  global container_id = 0
  global powder_id  = 0
  global bulk_density = 0
  global H          = 0
  global H_c          = 0
  global mouth_d     = 0
  global mouth_sh    = 0
  global length_c     = 0
  global diameter   = 0
  global empty_weight_g  = 0
  global volume_ml    = 0
  global shape_code   = 0
  global flow_code   = 0
  global shape = ""
  global Flowability = ""
  global full_weight_g = 0
  global cent_edge = 0
  global pick_2_base = 0.2 # distance from tcp to base of picking table
  global wall_thickness = 0.002

  def read_db_data():

    socket_open(SERVER_IP, SERVER_PORT)
    sleep(0.5)
    socket_send_string("GET_DATACODE_FLOATS")
    sleep(5)

    local fl = socket_read_ascii_float(14)
    socket_close()

    global container_id = fl[1]
    global powder_id = fl[2]
    global bulk_density = fl[3]
    global H          = fl[4]/1000
    global H_c          = fl[5]/1000
    global mouth_d     = fl[6]/1000
    global mouth_sh    = fl[7]/1000
    global length_c     = fl[8]/1000
    global diameter   = fl[9]/1000
    global empty_weight_g = fl[10]
    global volume_ml    = fl[11]
    global full_weight_g = fl[12]
    global flow_code   = fl[13]
    global shape_code   = fl[14]

  	if (flow_code == 1.0):
  	  global Flowability = "MEDIUM"
  	elif (flow_code == 2.0):
  	  global Flowability = "LOW"
  	else:
  	  global Flowability = "HIGH"
  	end

    if ( shape_code == 1.0):
  	shape = "cylindrical"
  	cent_edge =  diameter
    else:
  	shape = "cubical"
  	cent_edge =  length_c
    end

  end

  def send_picking_info(Pow_name, target_weight):
    socket_open(SERVER_IP, SERVER_PORT)
    cmd = "PICK:"+Pow_name+";"+to_str(target_weight)
    socket_send_string(cmd)
    sleep(0.1)
    socket_close()
  end

  #### POTS ####
  def tilt_send(angle):
  	socket_open(SERVER_IP, SERVER_PORT)
  	angle = 92.0 - angle
  	socket_send_string("TILT:"+to_str(angle))
  	sync()
  	sleep(0.5)
  	socket_close()
  end

  def CW_Rotate(angle):
  	socket_open(SERVER_IP, SERVER_PORT)
  	socket_send_string("CWROTATE:"+to_str(angle))
  	sync()
  	sleep(0.5)
  	socket_close()
  end

  def CCW_Rotate(angle):
  	socket_open(SERVER_IP, SERVER_PORT)
  	socket_send_string("CCWROTATE:"+to_str(angle))
  	sync()
  	sleep(0.5)
  	socket_close()
  end

  def CW_full_Rotate():
  	socket_open(SERVER_IP, SERVER_PORT)
  	socket_send_string("FULLROTATE:"+to_str(1))
  	sync()
  	sleep(0.5)
  	socket_close()
  end

  def CCW_full_Rotate():
  	socket_open(SERVER_IP, SERVER_PORT)
  	socket_send_string("FULLROTATE:"+to_str(-1))
  	sync()
  	sleep(0.5)
  	socket_close()
  end

  def tilt_to_home():
  	socket_open(SERVER_IP, SERVER_PORT)
  	socket_send_string("HOME")
  	sync()
  	sleep(0.5)
  	socket_close()
  end
  #######
  def vibration_1():
  	set_analog_out(0,0.4)
  	sleep(1)
  	set_analog_out(0,0.0)
  	sleep(0)
  end

  def vibration_2():
  	set_analog_out(0,0.4)
  	sleep(0.8)
  	set_analog_out(0,0.0)
  	sleep(0.2)
  end

  def vibration_3():
  	set_analog_out(0,0.4)
  	sleep(0.5)
  	set_analog_out(0,0.0)
  	sleep(0.3)
  end

  def vibration_4():
  	set_analog_out(0,0.4)
  	sleep(0.5)
  	set_analog_out(0, 0.0)
  	sleep(0.5)
  end

  def vibration_5():
  	set_analog_out(0,0.4)
  	sleep(0.2)
  	set_analog_out(0, 0.0)
  	sleep(0.8)
  end

  ##################

  global gear_2_holder = 0.018
  global gain_per_percent = 0.5
  global hinge_2_base = 0.0421
  global TCP_2_tip_x = 0.0047
  global spatula_len = 0.182
  global spatula_offset = p[TCP_2_tip_x,0,spatula_len,0,0,0]
  global SPATULA_L_VOL_ML = 5.0        # 1 teaspoon = 5 mL
  global SPATULA_M_VOL_ML = 1.25       # 1/4 teaspoon = 1.25 mL
  global SPATULA_S_VOL_ML = 0.15625    # 1/32 teaspoon = 0.15625 mL
  global SPATULA_FLAT_M_VOL_ML  = 2.2
  global SPATULA_FLAT_S_VOL_ML  = 0.7   #based on caluclations using rho = m/V

  def correction_reset():
  	global g_k = 0.0
  	global g_depth_corr = 0.0
  	global g_prev_cum_w = weight_value
  end

  def params_init():

  	global scoop_status= ""
  	global w_dosed_total = 0.0
  	global last_scale = 0.0
  	global tilt_angle_sent = 0.0
  	global level = 0.0
  	global target_g = 0.0
  	global angle_max = 70
  	global angle_min = 20
  	global ry_deg_safe = 0
  	global ry_deg = 0

  	global scoop_ct = 0
  	global error_sum = 0.0
  	global error_sq_sum = 0.0
  	global scoop_g = 0.0

  	global g_k =0.0
  	global g_eta = 0.3

  	global g_gain_scale = 0.07
  	global g_k_min = 0.0
  	global g_k_max = 0.09

  	# ---------- Damping ----------
  	global g_alpha_under = 0.75   # aggressive when undershooting
  	global g_alpha_over  = 0.30   # conservative when overshooting

  	# ---------- Search ----------
  	global g_engagement_min = 0.05
  	global g_search_step = 0.01      # 3 mm

  	# ---------- Deadband ----------
  	global g_tol = 0.02               # 20 mg minimum
  	global g_tol_ratio = 0.05         # ±5% of target

  	# ---------- Limits ----------
  	global g_corr_max = 0.020         # 20 mm maximum correction

  	# ---------- States ----------
  	global g_depth_corr = 0.0
  	global g_prev_cum_w = -1.0
  end

  def clamp(x, lo, hi):
  	if(x<lo):
  		return lo
  	elif (x>hi):
  		return hi
  	else:
  		return x
  	end
  end

  def compute_level_percent(W_now, weight_value):   # W_now = container+powder, weight_value = live scale reading
      global delta = weight_value - last_scale

      if (delta < 0.0):
          delta = 0.0
      end

      global w_dosed_total = w_dosed_total + delta
      global last_scale = weight_value     # update the last scale reading

      local W_eff = W_now - w_dosed_total
      if (W_eff <  empty_weight_g):
          W_eff =  empty_weight_g
      end

      # Compute powder level %
      level = 100.0 * (W_eff -  empty_weight_g) / (full_weight_g -  empty_weight_g)

      # Clamp to 0–100
      level = clamp(level, 0, 100)
    textmsg("deb 1 = ", level)
      return level
  end

  def deg2rad(d):
  	return d*3.141592/180
  end

  def my_abs(val):
  	if (val<0):
  		return -val
  	else:
  		return val
  	end
  end

  def compute_tilt_deg(level_percent):
  	angle = angle_min + gain_per_percent*(100.0-level_percent)

    	textmsg("deb 2 = ", angle)
  	return clamp(angle, angle_min, angle_max)
  end

  def tilt(level_percentage):
  	new_angle = compute_tilt_deg(level_percentage)
    	textmsg("deb angle 1 = ", new_angle)
  	global angle_rel = new_angle - tilt_angle_sent
    	textmsg("deb 2 = ", angle_rel)

  	if my_abs(angle_rel)>2.0:
    		textmsg("deb loop")
  		tilt_send(new_angle)
  		global angle_deg = new_angle
    		textmsg("deb 2 = ", angle_deg)
  		global tilt_angle_sent = new_angle
  		global p_center_vertical = center_pose()
  		global p_center = updated_center_pose(p_center_vertical, angle_deg)
  	end
    	textmsg("deb loop exit")

  	tilt_send(angle_deg)
    	textmsg("deb angle 2 =", angle_deg)

  end

  def compute_scoop_depth(level, weight_value, target_g):

      global scoop_depth_rel = ((100.0-level)/100.0)*(H-mouth_sh)

      if (g_prev_cum_w < 0):
          g_prev_cum_w = weight_value
          g_depth_corr = 0.0

      else:
          global scoop_g = weight_value - g_prev_cum_w
          g_prev_cum_w = weight_value

          local error = target_g - scoop_g
          local engagement = scoop_g / target_g

          local tol = g_tol_ratio * target_g
          if (tol < g_tol):
              tol = g_tol
          end
          if ((engagement < g_engagement_min) and (scoop_g < target_g)):
              g_depth_corr = g_depth_corr + g_search_step
          elif (my_abs(error) <= tol):
  			sync()
          else:
              local error_norm = my_abs(error / target_g)
              local g_target = clamp(g_gain_scale * error_norm,g_k_min,g_k_max)

              g_k = (1.0-g_eta) * g_k + g_eta * g_target
              if (error > 0):
                  local corr = g_k * error
                  g_depth_corr = g_depth_corr +g_alpha_under * corr
              else:
                  local corr = g_k * error
                  g_depth_corr = g_depth_corr +g_alpha_over * corr

              end
              g_depth_corr = clamp(g_depth_corr,-g_corr_max,g_corr_max)

          end
      end
      scoop_depth = scoop_depth_rel + g_depth_corr
      scoop_depth = clamp(scoop_depth, 0.0, H)
      return scoop_depth

  end

  def get_scoop_weight(spatula, bulk_density):

  	local vol = 0

  	if (spatula == "spatula_L"):
  		vol = SPATULA_L_VOL_ML
  		global spatula_depth = 0.015
  		global spatula_mid   = 0.016
  		global spatula_ry    = 0.0

  	elif (spatula == "spatula_M"):
  		vol = SPATULA_M_VOL_ML
  		global spatula_depth = 0.010
  		global spatula_mid   = 0.0105
  		global spatula_ry    = 0.0

  	elif (spatula == "spatula_S"):
  		vol = SPATULA_S_VOL_ML
  		global spatula_depth = 0.008
  		global spatula_mid   = 0.006
  		global spatula_ry    = 0.0

  	elif (spatula == "spatula_flat_M"):
  		vol = SPATULA_FLAT_M_VOL_ML
  		global spatula_depth = 0.005
  		global spatula_mid   = 0.02
  		global spatula_ry    = 4.0

  	elif (spatula == "spatula_flat_S"):
  		vol = SPATULA_FLAT_S_VOL_ML
  		global spatula_depth = 0.005
  		global spatula_mid   = 0.011
  		global spatula_ry    = 4.0
  	else:
  		textmsg("Unknown spatula type")
  		return 0.0
  	end
  	global target_g = vol * bulk_density
  	return target_g

  end

  def select_spatula(Flowability, level, diff, bulk_density, mouth_d ):

      local k = 1.1
      global powder_height = (H  - mouth_sh ) * level/100

      if (Flowability == "LOW"):
          local gFM = get_scoop_weight("spatula_flat_M", bulk_density)
  		local level_ok_FM = (mouth_d >= 0.05)
          local level_ok_FM = (spatula_mid  < powder_height)
          local diff_ok_FM  = (diff > k * gFM)
          local flatM_ok = level_ok_FM and diff_ok_FM
          if (flatM_ok):
              return "spatula_flat_M"
          else:
              return "spatula_flat_S"
          end
      end

      local gL = get_scoop_weight("spatula_L", bulk_density)
      local mouth_ok_L = (mouth_d  >= 0.05)
      local level_ok_L = (spatula_mid < powder_height)
      local diff_ok_L  = (diff > k * gL)

      local large_ok = mouth_ok_L and level_ok_L and diff_ok_L
      local gM = get_scoop_weight("spatula_M", bulk_density)
      local level_ok_M = (spatula_mid < powder_height)
      local diff_ok_M  = (diff > k * gM)

      local medium_ok = level_ok_M and diff_ok_M

      if (large_ok):
          return "spatula_L"
      elif (medium_ok):
          return "spatula_M"
      else:
          return "spatula_S"
      end
  end

  def after_scoop():
  	set_tcp(tcp_dosing)
  	set_analog_out(0,0.0)
  	tilt_send(angle_deg)
  	sleep(0.5)
  	movel(lifted_pose, a=0.05, v=0.2)
  	movel(tilted_pose_in_base2, a=0.05, v=0.2)
  	set_analog_out(0,0.4)
  	if (Flowability == "LOW"):
  		movel(end_rel_tilted_level2, a=0.03, v=0.1)
  		sleep(0.5)
  		movel(tilted_pose_in_base2, a=0.05, v=0.2)
  	  	movel(pose_trans(tilted_pose_in_base2, p[0,0,0,0,0,2.0]), a=0.05, v=0.2)
  		#movel(tilted_pose_in_base2, a=0.05, v=0.2)
  	else:
  	    movel(pose_trans(tilted_pose_in_base2, p[0,0,0,0,0,2.0]), a=0.05, v=0.2)
  	    movel(tilted_pose_in_base2, a=0.05, v=0.2)
  	end
  	set_analog_out(0,0.0)
  	movel(lifted_pose, a=0.5, v=0.5)
  	tilt_to_home()
  	set_tcp(tcp_default)
  end

  def center_pose():
  	global p_translated = container_place
  	#global p_translated = pots_axis_temp

  	#cx = p_translated[0]
  	#cy = p_translated[1]
  	#cz = p_translated[2]

  	global p_center_vertical_temp = pose_trans(p_translated, p[0,0,0, deg2rad(90), 0, 0])
  	cx = p_center_vertical_temp[0]
  	cy = p_center_vertical_temp[1]
  	cz = p_center_vertical_temp[2]
  	rx = p_center_vertical_temp[3]
  	ry = p_center_vertical_temp[4]
  	rz = p_center_vertical_temp[5]

  	global p_center_vertical_temp = p[cx,cy,cz, 0, 0, rz]
  	trans_rel = p[0,0,-pick_2_base+H,0,0,0]
  	global p_center_vertical =  pose_trans(p_center_vertical_temp, trans_rel)
  	return p_center_vertical
  end

  def updated_center_pose(p_center_vertical, angle_deg):
  	hinge_pose = pose_trans(p_center_vertical, p[0,0,-hinge_2_base-gear_2_holder-H ,0,0,0])
  	local_rel = pose_trans(pose_inv(hinge_pose), p_center_vertical)

  	rot_tilt = p[0,0,0, -deg2rad(angle_deg),0,0]
  	local_rel_tilted = pose_trans(rot_tilt, local_rel)

  	global p_center = pose_trans(hinge_pose, local_rel_tilted)
  	return p_center
  end

  def scoop_powder(p_center):
  	vibration_voltage = 0.4
  	global scoop_radius_default = 0.0

  	scoop_radius_default = mouth_d /2 - spatula_depth - wall_thickness
  	scoop_safe_entry_pose = pose_trans(p_center, p[-TCP_2_tip_x,0,spatula_len+0.05,0,0,0])
  	scoop_entry_pose = pose_trans(p_center, p[-TCP_2_tip_x,0,spatula_len,0,0,0])

  	movel(scoop_safe_entry_pose, a=0.1, v=0.25)
  	movel(scoop_entry_pose, a=0.1, v=0.25)

  	scoop_start_rel_int = p[0, 0, -mouth_sh , 0, 0, 0]
  	scoop_start_pose_int = pose_trans(scoop_entry_pose, scoop_start_rel_int)


  	#local ry_deg = map_tilt_to_ry_deg(angle_deg,level)
  	#local ry_result = map_tilt_to_ry_deg(angle_deg,level)

  	#global scoop_depth = compute_scoop_depth(level,weight_value, target_g)

  	global ry = deg2rad(90-angle_deg)

  	#global ry_safe = ry_result[0]
  	#global ry = deg2rad(ry_result[1])

  	if (spatula_mid < powder_height):

  		global total_depth = mouth_sh + scoop_depth + spatula_mid
  		global total_depth = clamp(total_depth, 0, H - spatula_mid)

  		safe_scoop_pivot = (mouth_d  - spatula_depth)/(total_depth)
  		global ry_safe = asin(safe_scoop_pivot)

  		scoop_start_rel = p[scoop_radius_default, 0, -total_depth, 0, 0, 0]

  		rot_mid = p[0, 0, 0, 0, 0, 0.785]
  		rot_end = p[0, 0, 0, 0, 0, 1.5708]

  		scoop_via_rel = pose_trans(rot_mid, scoop_start_rel)
  		scoop_end_rel = pose_trans(rot_end, scoop_start_rel)

  		scoop_start_pose = pose_trans(scoop_entry_pose, scoop_start_rel)
  		scoop_via_pose = pose_trans(scoop_entry_pose, scoop_via_rel)
  		scoop_end_pose = pose_trans(scoop_entry_pose, scoop_end_rel)


  			if (Flowability == "LOW"):
  				movel(pose_trans(scoop_start_pose_int,p[0,0,0,0,0,-1.5708]), a=0.1, v=0.25)
  				local spatula_base = pose_trans(scoop_entry_pose, p[0, 0, -H+wall_thickness, 0, 0, 0])
  				local scrape_pivot = pose_trans(scoop_entry_pose, p[0,0, -spatula_len,0,0,0])

  				global sticky_in_angle = -atan((cent_edge/2-spatula_depth)/H)
  				spatula_tilt_rel = pose_trans(pose_inv(scrape_pivot), spatula_base)

  				spatula_tilt = pose_trans(spatula_tilt_rel, p[0, 0, 0, 0, sticky_in_angle, 0])
  				global tilted_pose = pose_trans(scrape_pivot, p[0,0,0,spatula_tilt[3],spatula_tilt[4], spatula_tilt[5]])

  				global tilted_pose = pose_trans(tilted_pose, p[0,0,spatula_len-H+wall_thickness,0,0,0])
  				global rotate_90=pose_trans(tilted_pose,p[0,0,0,0,0,-1.5708])


  				movel(rotate_90,a=0.1, v=0.25)

  				#global sticky_in_angle = -atan((cent_edge/2-wall_thickness-spatula_depth)/(total_depth+spatula_mid))
  				#local scrape_target = pose_trans(scoop_entry_pose, p[0,0,-total_depth-spatula_mid,0,0,0])
  				#local scrape_pivot = pose_trans(scoop_entry_pose, p[0,0,-spatula_len,0,0,0])
  				#local scrape_rel = pose_trans(pose_inv(scrape_pivot), scrape_target)
  				#local scoop_sticky_in = pose_trans(scrape_rel, p[0,0,0,0,sticky_in_angle,0])

  				#global scrape_pose = pose_trans(scrape_pivot, p[0,0,0,scoop_sticky_in[3],scoop_sticky_in[4], scoop_sticky_in[5]])
  				#global scrape_pose = pose_trans(scrape_pose, p[0,0,spatula_len-total_depth-spatula_mid,0,0,0])

  				#scoop_sticky_in = pose_trans(scoop_start_pose, p[0,0,0,0,sticky_in_angle,0])
  				#movel(scrape_pose, a=0.1, v=0.25)
  				#movel(scrape_target,a=0.1,v=0.25)
  				CW_full_Rotate()
  				movel(scoop_start_pose, a=0.1, v=0.25)

  			else:
  				movel(scoop_start_pose_int, a=0.1, v=0.25)
  				movel(scoop_start_pose, a=0.1, v=0.25)
  				CW_full_Rotate()
  			end

  		movec(scoop_via_pose, scoop_end_pose, a=0.05, v=0.04)
  		#sleep(1.0)

  		# safe_retention
  		local pivot_pose = pose_trans(scoop_end_pose, p[0,0,total_depth-spatula_len,0,0,0])
  		local end_rel = pose_trans(pose_inv(pivot_pose), scoop_end_pose)
  		local end_rel_tilted = pose_trans(end_rel, p[0, 0, 0, 0, ry_safe-deg2rad(spatula_ry), 0])
  		local tilted_pose_in_base = pose_trans(pivot_pose, p[0,0,0,end_rel_tilted[3],end_rel_tilted[4], end_rel_tilted[5]])
  		local tilted_pose_in_base = pose_trans(tilted_pose_in_base, p[0, 0, spatula_len-total_depth, 0, 0, 0])
  		# sptula pivoted around the container rim of the mouth at ry_safe
  		movel(tilted_pose_in_base, a=0.03, v=0.1)

  		global safe_x = sin(ry_safe)*(total_depth-mouth_sh - (mouth_d - spatula_depth)*tan(ry_safe/2))
  		global safe_z = cos(ry_safe)*(total_depth-mouth_sh - (mouth_d - spatula_depth)*tan(ry_safe/2))

  		local safe_up = pose_trans(tilted_pose_in_base, p[-safe_x,0,safe_z,0,0,0])
  		movel(safe_up, a=0.03, v=0.1)

  		# full exit
  		local pivot_pose2 = pose_trans(scoop_entry_pose, p[0,0,-spatula_len,0,0,0])
  		local end_rel2 = pose_trans(pose_inv(pivot_pose2), tilted_pose_in_base)
  		#popup("is the spatula crashing front? ", blocking = True)
  		local end_rel_tilted2 = pose_trans(end_rel2, p[0, 0, 0, 0, ry-ry_safe-deg2rad(spatula_ry), 0])

  	else : # emptying logic
  		CCW_full_Rotate()

  		spatula_base = pose_trans(scoop_entry_pose, p[0, 0, -H+wall_thickness, 0, 0, 0])
  		local pivot_pose2 = pose_trans(scoop_entry_pose, p[0,0,-spatula_len,0,0,0])
  		# tilt inwards
  		global in_angle = -atan((cent_edge/2-spatula_depth)/H)
  		spatula_tilt_rel = pose_trans(pose_inv(pivot_pose2), spatula_base)

  		spatula_tilt = pose_trans(spatula_tilt_rel, p[0, 0, 0, -in_angle, 0, 0])
  		global tilted_pose = pose_trans(pivot_pose2, p[0,0,0,spatula_tilt[3],spatula_tilt[4], spatula_tilt[5]])

  		global tilted_pose = pose_trans(tilted_pose, p[0,0,spatula_len-H+wall_thickness,0,0,0])

  		movel(tilted_pose,a=0.1, v=0.25)

  		rotate90=pose_trans(tilted_pose,p[0,0,0,0,0,1.5708])

  		#sleep(1)
  		#Rotate()
  		#sleep(0.2)
  		movel(rotate90, a=0.1, v=0.1)
  		#popup("is the spatula crashing front? ", blocking = True)
  		movel(pose_trans(scoop_start_pose_int,p[0,0,0,0,0,1.5708]), a=0.03, v=0.1)
  		# full exit
  		#local pivot_pose2 = pose_trans(scoop_entry_pose, p[0,0,-spatula_len,0,0,0])
  		local end_rel2 = pose_trans(pose_inv(scoop_entry_pose), rotate90)
  		local end_rel_tilted2 = pose_trans(end_rel2, p[0, 0, 0, 0, ry-in_angle-deg2rad(spatula_ry), 0])
  	end

  	# exit flat spoon
  	global tilted_pose_in_base2 = pose_trans(pivot_pose2, p[0,0,0,end_rel_tilted2[3],end_rel_tilted2[4], end_rel_tilted2[5]])
  	global tilted_pose_in_base2 = pose_trans(tilted_pose_in_base2, p[0, 0, spatula_len-spatula_mid, 0, 0, 0])
  	# spaula exited at center of the mouth at ry
  	movel(tilted_pose_in_base2, a=0.03, v=0.1)
  	if(scoop_status== "normal"):
  		vib_thread=True
  		if (spatula=="spatula_S"):
  			vibration_3()
  			local ry_level = deg2rad(12)
  		elif(spatula=="spatula_flat_S" or spatula=="spatula_flat_M"):
  			vibration_3()
  			local ry_level = deg2rad(5)
  		else:
  			set_analog_out(0,0.4)
  			local ry_level = deg2rad(25)
  		end

  		# remove excess
  		local pivot_pose_level = pose_trans(tilted_pose_in_base2, p[0,0,-spatula_len,0,0,0])
  		local end_rel_level = pose_trans(pose_inv(pivot_pose_level), tilted_pose_in_base2)
  		local end_rel_tilted_level = pose_trans(end_rel_level, p[0, 0, 0, 0, -ry_level, 0])
  		global end_rel_tilted_level2 = pose_trans(pivot_pose_level, p[0, 0, 0,end_rel_tilted_level[3],end_rel_tilted_level[4], end_rel_tilted_level[5]])
  		global end_rel_tilted_level2 = pose_trans(end_rel_tilted_level2, p[0,0,spatula_len,0,0,0])
  		movel(end_rel_tilted_level2, a=0.03, v=0.1)

  		if (spatula == "spatula_flat_S" or spatula == "spatula_flat_M"):
  			vib_thread=False
  			set_analog_out(0, 0.0)
  		end
  	else:
  		set_analog_out(0, 0.0)
  	end
  	movel(tilted_pose_in_base2, a=0.03, v=0.1)
  	set_analog_out(0, 0.0)
  	vib_thread=False
  	global lifted_pose = pose_trans(tilted_pose_in_base2, p[-0.04,0,0.04,0,0,0]) # safety distance away from the container

  	movel(lifted_pose, a=0.03, v=0.1)
  	tilt_to_home()
  end

  def auto_tilt_and_scoop(W_now, target_weight, weight_value):
  	set_tcp(tcp_dosing)
  	global level = compute_level_percent(W_now, weight_value)

  	global spatula = select_spatula(Flowability, level, diff, bulk_density, mouth_d )
  	textmsg("deb 4 = ", spatula)
  	global target_g = get_scoop_weight(spatula, bulk_density)
  	textmsg("deb 5 = ", target_g)

  	global scoop_depth = compute_scoop_depth(level, weight_value, target_g)
    	textmsg("deb 6 = ", scoop_depth)
  	tilt(level)

  	scoop_powder(p_center)

  	#textmsg("deb 7 - sucess")
   	set_tcp(tcp_default)
  end
  $ 21 "Script: Weight_scale_socket_s.script"
  global s_depth = 0
  global s_length =0
  global s_volume = 0
  global ry_theta  = 0

  def get_weight():
  	socket_open(SERVER_IP,SERVER_PORT)
  	#sleep(0.2)
  	textmsg("socket opened successfully!")
  	socket_send_string("GET_WEIGHT")
  	#sleep(0.2)
  	sync()
  	receiveFromServ = socket_read_ascii_float(1)
  	#sleep(1)
  	while (receiveFromServ[0] < 1):
  		receiveFromServ = socket_read_ascii_float(1)
  		sleep(0.01)
  	end
  	textmsg("Received weight:", receiveFromServ[1])
  	#sleep(0.2)
  	socket_close()
  	#sleep(0.2)
  	return receiveFromServ[1]
  end

  def tare_scale():
  	socket_open(SERVER_IP,SERVER_PORT)
  	socket_send_string("TARE")
  	sleep(2)
  	socket_close()
  end

  def zero_scale():
  	socket_open(SERVER_IP,SERVER_PORT)
  	socket_send_string("ZERO")
  	sleep(0.5)
  	socket_close()
  end

  def log_weight():
  	socket_open(SERVER_IP,SERVER_PORT)
  	socket_send_string("LOG_WEIGHT")
  	sleep(0.5)
  	socket_close()
  end

  def send_target_info():
  	socket_open(SERVER_IP,SERVER_PORT)
  	socket_send_string("SET_TARGET:" + to_str(target_weight))
  	sleep(0.2)
  	socket_close()
  end
  def send_powder_info():
  	socket_open(SERVER_IP,SERVER_PORT)
  	socket_send_string("SET_POWDER:" + Pow_name)
  	sleep(0.2)
  	socket_close()
  end
  def send_spatula_info():
  	socket_open(SERVER_IP,SERVER_PORT)
  	socket_send_string("SET_SPATULA:" + spatula)
  	#sleep(1)

  	#local fl = socket_read_ascii_float(4)

    	#global s_depth = fl[1]
    	#global s_length = fl[2]
   	#global s_volume = fl[3]
   	#global ry_theta  = fl[4]
  	sleep(0.2)
  	socket_close()
  end

  def send_level_info():
  	socket_open(SERVER_IP,SERVER_PORT)
  	socket_send_string("SET_LEVEL:" + to_str(level))
  	sleep(0.2)
  	socket_close()
  end

  def get_cont_weight():
    socket_open(SERVER_IP, SERVER_PORT)
    #rq_open_and_wait()
    cmd = "GET_CONT_WEIGHT"
    socket_send_string(cmd)
    sync()
    sleep(0.5)
    receiveFromSer = socket_read_ascii_float(1)
    socket_close()
    return receiveFromSer[1]
  end

  $ 22 "BeforeStarts"
  $ 23 "uLM"
  $ 24 "CMD_Stop≔ False "
  global CMD_Stop=  False
  $ 25 "CMD_Abort≔ False "
  global CMD_Abort=  False
  $ 26 "CMD_Clear≔ False "
  global CMD_Clear=  False
  $ 27 "STATE≔1"
  global STATE=1
  $ 28 "STATE_Info≔''"
  global STATE_Info=""
  $ 29 "ARM_Referenced≔ False "
  global ARM_Referenced=  False
  $ 30 "zero_ftsensor()"
  zero_ftsensor()
  $ 31 "poses init"
  $ 32 "PSE_A≔p[0,0,0,0,0,0]"
  global PSE_A=p[0,0,0,0,0,0]
  $ 33 "PSE_A_H≔p[0,0,0,0,0,0]"
  global PSE_A_H=p[0,0,0,0,0,0]
  $ 34 "PSE_R≔p[0,0,0,0,0,0]"
  global PSE_R=p[0,0,0,0,0,0]
  $ 35 "PSE_R_H≔p[0,0,0,0,0,0]"
  global PSE_R_H=p[0,0,0,0,0,0]
  $ 36 "PSE_T≔p[0,0,0,0,0,0]"
  global PSE_T=p[0,0,0,0,0,0]
  $ 37 "PSE_T_H≔p[0,0,0,0,0,0]"
  global PSE_T_H=p[0,0,0,0,0,0]
  $ 38 "PSE_C_E≔p[0,0,0,0,0,0]"
  global PSE_C_E=p[0,0,0,0,0,0]
  $ 39 "PSE_C_H≔p[0,0,0,0,0,0]"
  global PSE_C_H=p[0,0,0,0,0,0]
  $ 40 "PSE_C_S≔p[0,0,0,0,0,0]"
  global PSE_C_S=p[0,0,0,0,0,0]
  $ 41 "init_home_by_cartesian_pose(p[0,-0.400,0.300,0,0,0])"
  init_home_by_cartesian_pose(p[0,-0.400,0.300,0,0,0])
  $ 42 "Clearing"
  $ 43 "reset_error()"
  reset_error()
  $ 44 "reset_warning()"
  reset_warning()
  $ 45 "uGo"
  $ 47 "ugo_init( True ,'http://192.168.12.120:10001')"
  ugo_init(  True  ,"http://192.168.12.120:10001")
  $ 48 "ugo_update_outputs()"
  ugo_update_outputs()
  $ 49 "App"
  $ 50 "'ADD APPLICATION SPECIFIC COMMANDS'"
  # 'ADD APPLICATION SPECIFIC COMMANDS'
  $ 51 "Tools"
  $ 52 "OBJ_Picked≔gripper_has_object()"
  global OBJ_Picked=gripper_has_object()
  $ 53 "If OBJ_Picked"
  if (OBJ_Picked):
    # begin: URCap Program Node
    #   Source: Robotiq_Grippers, 3.17.0.105337, Robotiq Inc.
    #   Type: Gripper Activate
    $ 54 "Gripper Activate"

    kill rq_gripper_communication_thread
    rq_gripper_communication_thread_started = False
    rq_close_gripper_socket("1")
    rq_close_gripper_socket("2")
    rq_close_gripper_socket("3")
    rq_close_gripper_socket("4")

    rq_init_comm_if_connected(9, "1")
    rq_init_comm_if_connected(2, "2")
    rq_init_comm_if_connected(3, "3")
    rq_init_comm_if_connected(4, "4")
    rq_print_connected_grippers()
    rq_gripper_communication_thread = run rq_gripper_communication()

    while(not rq_gripper_communication_thread_started):
        sleep(0.008)
    end

    rq_set_max_current_for_all_grippers()

    reset_and_activate = False

    rq_activate_all_grippers(False)
    # end: URCap Program Node
  else:
    $ 55 "Else" "noBreak"
    # begin: URCap Program Node
    #   Source: Robotiq_Grippers, 3.17.0.105337, Robotiq Inc.
    #   Type: Gripper Activate
    $ 56 "Gripper Reset and Activate"

    kill rq_gripper_communication_thread
    rq_gripper_communication_thread_started = False
    rq_close_gripper_socket("1")
    rq_close_gripper_socket("2")
    rq_close_gripper_socket("3")
    rq_close_gripper_socket("4")

    rq_init_comm_if_connected(9, "1")
    rq_init_comm_if_connected(2, "2")
    rq_init_comm_if_connected(3, "3")
    rq_init_comm_if_connected(4, "4")
    rq_print_connected_grippers()
    rq_gripper_communication_thread = run rq_gripper_communication()

    while(not rq_gripper_communication_thread_started):
        sleep(0.008)
    end

    rq_set_max_current_for_all_grippers()

    reset_and_activate = True

    rq_activate_all_grippers(True)
    # end: URCap Program Node
  end
  $ 57 "zero_ftsensor()"
  zero_ftsensor()
  $ 58 "EXTT"
  $ 59 "Set GRP_3F_Enable=Off"
  set_standard_digital_out(4, False)
  $ 60 "Set BarcodeTrigger=Off"
  set_standard_digital_out(6, False)
  $ 61 "Set GRP_3F_Decap=Off"
  set_standard_digital_out(3, False)
  $ 62 "Set GRP_3F_Cap=Off"
  set_standard_digital_out(2, False)
  $ 63 "Set GRP_3F_Open=Off"
  set_standard_digital_out(5, False)
  $ 64 "PSE_T≔get_tool_free_pose(dir=[0,0,0.150], move_in_base_frame=True)"
  global PSE_T=get_tool_free_pose(dir=[0,0,0.150], move_in_base_frame=True)
  $ 65 "If is_reachable(Base_const, [PSE_T])"
  if (is_reachable(p[0.0,0.0,0.0,0.0,0.0,0.0], [PSE_T])):
    $ 66 "MoveL"
    $ 67 "PSE_T" "breakAfter"
    movel(PSE_T, a=1.2, v=0.15)
  end
  $ 68 "powder dispensing variable init"
  $ 69 "Start_thread≔ False "
  global Start_thread=  False
  $ 70 "vib_thread≔ False "
  global vib_thread=  False
  $ 71 "w_full_thread≔ False "
  global w_full_thread=  False
  $ 72 "Picking≔ False "
  global Picking=  False
  $ 73 "d_cc≔0.07"
  global d_cc=0.07
  $ 74 "kp≔0.0035"
  global kp=0.0035
  $ 75 "ki≔0.0001"
  global ki=0.0001
  $ 76 "kd≔0.003"
  global kd=0.003
  $ 77 "dt≔0.2"
  global dt=0.2
  $ 78 "Integral_error≔0"
  global Integral_error=0
  $ 79 "current_error≔0"
  global current_error=0
  $ 80 "previous_error≔0"
  global previous_error=0
  $ 81 "tilt_increment≔0"
  global tilt_increment=0
  $ 82 "tilt_angle≔0"
  global tilt_angle=0
  $ 83 "diff≔0"
  global diff=0
  $ 84 "tilt_to_home()"
  tilt_to_home()
  $ 85 "params_init()"
  params_init()
  $ 86 "switch_spat_M≔ True "
  global switch_spat_M=  True
  $ 87 "switch_spat_S≔ True "
  global switch_spat_S=  True
  $ 88 "switch_spat_F_M≔ True "
  global switch_spat_F_M=  True
  $ 89 "switch_spat_F_S≔ True "
  global switch_spat_F_S=  True
  $ 90 "last_scale≔0"
  global last_scale=0
  $ 843 "Thread_1"
  thread Thread_1():
    while (True):
      $ 844 "Dosing Weight"
      $ 845 "If Start_thread≟ True "
      if (Start_thread ==   True  ):
        $ 846 "weight_value≔get_weight()"
        global weight_value=get_weight()
        $ 847 "diff≔target_weight-weight_value"
        global diff=target_weight-weight_value
        $ 848 "Wait: 0.2"
        sleep(0.2)
        $ 849 "sync()"
        sync()
      end
      $ 850 "sync()"
      sync()
    end
  end
  threadId_Thread_1 = run Thread_1()
  $ 851 "Thread_2"
  thread Thread_2():
    while (True):
      $ 852 "Vibration motor"
      $ 853 "Loop vib_thread≟ True "
      thread Thread_while_853():
        while (True):
          $ 854 "diff≔target_weight-weight_value"
          global diff=target_weight-weight_value
          $ 855 "If diff>0.02 and spatula≠'spatula_flat_S' "
          global thread_flag_855=0
          thread Thread_if_855():
            $ 857 "Set AO[0]=4.0"
            set_standard_analog_out(0, 0.4)
            thread_flag_855 = 1
          end
          if (diff>0.02  and  spatula != "spatula_flat_S" ):
            global thread_handler_855=run Thread_if_855()
            while (thread_flag_855 == 0):
              if not(diff>0.02  and  spatula != "spatula_flat_S" ):
                kill thread_handler_855
                thread_flag_855 = 2
              else:
                sync()
              end
            end
          else:
            thread_flag_855 = 2
          end
          if (thread_flag_855 == 2):
            $ 858 "ElseIf diff>0.02 and spatula≟'spatula_flat_S'"
            if (diff>0.02 and spatula == "spatula_flat_S"):
              $ 859 "vibration_3()"
              vibration_3()
            else:
              $ 860 "ElseIf diff≤0.03"
              global thread_flag_860=0
              thread Thread_if_860():
                $ 861 "vibration_2()"
                vibration_2()
                thread_flag_860 = 1
              end
              if (diff <= 0.03):
                global thread_handler_860=run Thread_if_860()
                while (thread_flag_860 == 0):
                  if not(diff <= 0.03):
                    kill thread_handler_860
                    thread_flag_860 = 2
                  else:
                    sync()
                  end
                end
              else:
                thread_flag_860 = 2
              end
              if (thread_flag_860 == 2):
                $ 862 "Else" "noBreak"
                $ 863 "Set AO[0]=0.0"
                set_standard_analog_out(0, 0.0)
              end
            end
          end
        end
      end
      if (vib_thread ==   True  ):
        global thread_handler_853=run Thread_while_853()
        while (vib_thread ==   True  ):
          sync()
        end
        kill thread_handler_853
      end
      $ 864 "sync()"
      sync()
    end
  end
  threadId_Thread_2 = run Thread_2()
  $ 865 "Thread_3"
  thread Thread_3():
    while (True):
      $ 866 "Container weight"
      $ 867 "If w_full_thread≟ True "
      if (w_full_thread ==   True  ):
        $ 868 "aa_weight_cont≔get_cont_weight()"
        global aa_weight_cont=get_cont_weight()
        $ 869 "Wait: 0.2"
        sleep(0.2)
        $ 870 "sync()"
        sync()
      end
      $ 871 "sync()"
      sync()
    end
  end
  threadId_Thread_3 = run Thread_3()
  while (True):
    $ 91 "Robot Program"
    $ 92 "MAIN"
    $ 93 "command_manager(external_control='uGO', cond_suspend=(ITM_Manipulated and AMR_AtTarget and AMR_Charging and AMR_Battery<40), cond_unsuspend=(AMR_Battery≟60))"
    command_manager(external_control="uGO", cond_suspend=(ITM_Manipulated  and  AMR_AtTarget  and  AMR_Charging  and  AMR_Battery<40), cond_unsuspend=(AMR_Battery == 60))
    $ 94 "log_state(STATE_Info)"
    log_state(STATE_Info)
    $ 95 "Switch STATE"
    switch_1 = STATE
    $ 96 "Case 1"
    if (1 == switch_1):
      $ 97 "Stopping"
      $ 98 "STATE_Info≔'Stopping'"
      global STATE_Info="Stopping"
      $ 99 "end_freedrive_mode()"
      end_freedrive_mode()
      $ 100 "Set"
      set_tcp(p[0.0,0.0,0.161,3.1415,0.0,0.0])
      $ 101 "PSE_T≔get_tool_free_pose(dir=[0,0,0.150], move_in_base_frame=True)"
      global PSE_T=get_tool_free_pose(dir=[0,0,0.150], move_in_base_frame=True)
      $ 102 "If is_reachable(Base_const, [PSE_T])"
      if (is_reachable(p[0.0,0.0,0.0,0.0,0.0,0.0], [PSE_T])):
        $ 103 "MoveL"
        $ 104 "PSE_T" "breakAfter"
        movel(PSE_T, a=1.2, v=0.15)
      end
      $ 105 "do_transition(keep_rxry=OBJ_Picked, r=0)"
      do_transition(keep_rxry=OBJ_Picked, r=0)
      $ 114 "Call Sub_AMR_MiR_V3"
      Sub_AMR_MiR_V3()
      $ 115 "If stopping() and AMR_Done"
      if (stopping()  and  AMR_Done):
        $ 116 "STATE≔2"
        global STATE=2
        $ 117 "ugo_update_outputs()"
        ugo_update_outputs()
      end
    elif (2 == switch_1):
      $ 118 "Case 2"
      $ 119 "Stopped"
      $ 120 "STATE_Info≔'Stopped'"
      global STATE_Info="Stopped"
      $ 121 "Call Sub_AMR_MiR_V3"
      Sub_AMR_MiR_V3()
      $ 122 "If CMD_Reset  or PB_Start"
      if (CMD_Reset   or  get_standard_digital_in(0)):
        $ 123 "STATE≔3"
        global STATE=3
        $ 124 "ugo_update_outputs()"
        ugo_update_outputs()
      end
    elif (3 == switch_1):
      $ 125 "Case 3"
      $ 126 " Resetting"
      $ 127 "STATE_Info≔'Resetting'"
      global STATE_Info="Resetting"
      $ 128 "uML"
      $ 129 "reset_error()"
      reset_error()
      $ 130 "reset_warning()"
      reset_warning()
      $ 131 "PROCESS_Step≔0"
      global PROCESS_Step=0
      $ 132 "PROCESS_Info≔''"
      global PROCESS_Info=""
      $ 133 "ARM_Referenced≔ False "
      global ARM_Referenced=  False
      $ 134 "WRK_Done≔ False "
      global WRK_Done=  False
      $ 135 "ITM_Prepared≔ False "
      global ITM_Prepared=  False
      $ 136 "ITM_Manipulated≔ False "
      global ITM_Manipulated=  False
      $ 137 "STP≔0"
      global STP=0
      $ 138 "Action≔0"
      global Action=0
      $ 139 "Action_Info≔''"
      global Action_Info=""
      $ 140 "ITM_ID≔0"
      global ITM_ID=0
      $ 141 "JIG≔0"
      global JIG=0
      $ 142 "JIG_Slot≔0"
      global JIG_Slot=0
      $ 143 "Task_info≔''"
      global Task_info=""
      $ 144 "Set"
      set_tcp(p[0.0,0.0,0.161,3.1415,0.0,0.0])
      $ 145 "App"
      $ 146 "'ADD APPLICATION SPECIFIC COMMANDS'"
      # 'ADD APPLICATION SPECIFIC COMMANDS'
      $ 147 "OBJ_Type≔0"
      global OBJ_Type=0
      $ 148 "OBJ_Nbr≔0"
      global OBJ_Nbr=0
      $ 149 "If CNT_Rack_Output≥50"
      if (CNT_Rack_Output >= 50):
        $ 150 "CNT_Rack_Output≔0"
        global CNT_Rack_Output=0
      end
      $ 151 "TASK≔struct(ID=0, NAVI=struct(target=0, footprint=0, protectiveOff=0, dock=0), WORK=struct(ITM_ID_Src=0, JIG_ID_Src=0, OBJ_Nbr_Src=0, ACT_Src=0, ITM_ID_Tgt=0, JIG_ID_Tgt=0, OBJ_Nbr_Tgt=0, ACT_Tgt=0, OBJ_Type=0))"
      global TASK=struct(ID=0, NAVI=struct(target=0, footprint=0, protectiveOff=0, dock=0), WORK=struct(ITM_ID_Src=0, JIG_ID_Src=0, OBJ_Nbr_Src=0, ACT_Src=0, ITM_ID_Tgt=0, JIG_ID_Tgt=0, OBJ_Nbr_Tgt=0, ACT_Tgt=0, OBJ_Type=0))
      $ 152 "Call Sub_AMR_MiR_V3"
      Sub_AMR_MiR_V3()
      $ 153 "If resetting() and AMR_Done"
      if (resetting()  and  AMR_Done):
        $ 154 "STATE≔4"
        global STATE=4
        $ 155 "ugo_update_outputs()"
        ugo_update_outputs()
      end
    elif (4 == switch_1):
      $ 156 "Case 4"
      $ 157 "Idle"
      $ 158 "STATE_Info≔'Idle'"
      global STATE_Info="Idle"
      $ 159 "If CMD_Start"
      if (CMD_Start):
        $ 160 "STATE≔5"
        global STATE=5
        $ 161 "ugo_update_outputs()"
        ugo_update_outputs()
      end
    elif (5 == switch_1):
      $ 162 "Case 5"
      $ 163 "Starting"
      $ 164 "STATE_Info≔'Starting'"
      global STATE_Info="Starting"
      $ 165 "'ADD COMMANDS WHAT TO START WITH'"
      # 'ADD COMMANDS WHAT TO START WITH'
      $ 166 "Call Sub_AMR_MiR_V3"
      Sub_AMR_MiR_V3()
      $ 167 "get ugo data"
      $ 168 "Assign Tasks"
      $ 169 "TASK.ID = ugo_get_task()"
      TASK.ID = ugo_get_task()
      $ 170 "If TASK.ID≟1"
      if (TASK.ID == 1):
        $ 171 "Task_info≔'Charge'"
        global Task_info="Charge"
        $ 172 "Parameters"
        $ 173 "AMR_PosTarget≔1"
        global AMR_PosTarget=1
      else:
        $ 174 "ElseIf TASK.ID≟9"
        if (TASK.ID == 9):
          $ 175 "'Pick Sarstedt Rack from Variable source'"
          # 'Pick Sarstedt Rack from Variable source'
          $ 176 "Task_info≔'Navigate to Target'"
          global Task_info="Navigate to Target"
          $ 177 "Parameters"
          $ 178 "AMR_PosTarget≔UGO.read_input('00','ITM_ID')"
          global AMR_PosTarget=UGO.read_input("00","ITM_ID")
        else:
          $ 179 "ElseIf TASK.ID≟13"
          if (TASK.ID == 13):
            $ 180 "Task_info≔'Dose Powder'"
            global Task_info="Dose Powder"
            $ 181 "Parameters"
            $ 182 "ITM_ID≔1"
            global ITM_ID=1
            $ 183 "W_now≔(UGO.read_input('00','Container_weight'))/1000"
            global W_now=(UGO.read_input("00","Container_weight"))/1000
            $ 184 "Pow_name≔(UGO.read_input('00','Powder_name'))"
            global Pow_name=(UGO.read_input("00","Powder_name"))
            $ 185 "target_weight≔(UGO.read_input('00','Target_weight'))/1000"
            global target_weight=(UGO.read_input("00","Target_weight"))/1000
            $ 186 "params_init()"
            params_init()
            $ 187 "send_picking_info(Pow_name,target_weight)"
            send_picking_info(Pow_name,target_weight)
            $ 189 "OBJ_Type≔6"
            global OBJ_Type=6
            $ 190 "JIG≔17"
            global JIG=17
            $ 191 "AMR_PosTarget≔5"
            global AMR_PosTarget=5
          else:
            $ 192 "ElseIf TASK.ID≟49"
            if (TASK.ID == 49):
              $ 193 "Task_info≔'Pick Containers'"
              global Task_info="Pick Containers"
              $ 194 "Parameters"
              $ 195 "ITM_ID≔1"
              global ITM_ID=1
              $ 196 "OBJ_Type≔6"
              global OBJ_Type=6
              $ 197 "JIG≔15"
              global JIG=15
              $ 198 "AMR_PosTarget≔3"
              global AMR_PosTarget=3
            else:
              $ 199 "ElseIf TASK.ID≟50"
              if (TASK.ID == 50):
                $ 200 "Task_info≔'Decap Containers'"
                global Task_info="Decap Containers"
                $ 201 "Parameters"
                $ 202 "ITM_ID≔1"
                global ITM_ID=1
                $ 203 "OBJ_Type≔6"
                global OBJ_Type=6
                $ 204 "JIG≔16"
                global JIG=16
                $ 205 "AMR_PosTarget≔5"
                global AMR_PosTarget=5
              else:
                $ 206 "ElseIf TASK.ID≟51"
                if (TASK.ID == 51):
                  $ 207 "Task_info≔'Detect Spatula and transfer powder'"
                  global Task_info="Detect Spatula and transfer powder"
                  $ 208 "Parameters"
                  $ 209 "ITM_ID≔1"
                  global ITM_ID=1
                  $ 210 "target_weight≔(UGO.read_input('00','Target_weight'))/1000"
                  global target_weight=(UGO.read_input("00","Target_weight"))/1000
                  $ 211 "OBJ_Type≔8"
                  global OBJ_Type=8
                  $ 212 "JIG≔16"
                  global JIG=16
                  $ 213 "AMR_PosTarget≔5"
                  global AMR_PosTarget=5
                else:
                  $ 214 "ElseIf TASK.ID≟52"
                  if (TASK.ID == 52):
                    $ 215 "Task_info≔'Pick Powder'"
                    global Task_info="Pick Powder"
                    $ 216 "Parameters"
                    $ 217 "ITM_ID≔1"
                    global ITM_ID=1
                    $ 219 "OBJ_Type≔6"
                    global OBJ_Type=6
                    $ 220 "JIG≔15"
                    global JIG=15
                    $ 221 "AMR_PosTarget≔3"
                    global AMR_PosTarget=3
                  else:
                    $ 222 "ElseIf TASK.ID≟53"
                    if (TASK.ID == 53):
                      $ 223 "Task_info≔'Decap Powder'"
                      global Task_info="Decap Powder"
                      $ 224 "Parameters"
                      $ 225 "ITM_ID≔1"
                      global ITM_ID=1
                      $ 226 "OBJ_Type≔6"
                      global OBJ_Type=6
                      $ 227 "JIG≔1"
                      global JIG=1
                      $ 228 "AMR_PosTarget≔5"
                      global AMR_PosTarget=5
                    else:
                      $ 229 "ElseIf TASK.ID≟54"
                      if (TASK.ID == 54):
                        $ 230 "Task_info≔'Empty and swap Powder container'"
                        global Task_info="Empty and swap Powder container"
                        $ 239 "Parameters"
                        $ 240 "ITM_ID≔1"
                        global ITM_ID=1
                        $ 242 "W_now≔(UGO.read_input('00','Container_weight'))/1000"
                        global W_now=(UGO.read_input("00","Container_weight"))/1000
                        $ 243 "Pow_name≔(UGO.read_input('00','Powder_name'))"
                        global Pow_name=(UGO.read_input("00","Powder_name"))
                        $ 246 "OBJ_Type≔6"
                        global OBJ_Type=6
                        $ 247 "JIG≔17"
                        global JIG=17
                        $ 248 "AMR_PosTarget≔5"
                        global AMR_PosTarget=5
                      else:
                        $ 249 "ElseIf TASK.ID≟55"
                        if (TASK.ID == 55):
                          $ 250 "Task_info≔'Place Powder'"
                          global Task_info="Place Powder"
                          $ 251 "Parameters"
                          $ 252 "ITM_ID≔1"
                          global ITM_ID=1
                          $ 253 "OBJ_Type≔6"
                          global OBJ_Type=6
                          $ 254 "JIG≔21"
                          global JIG=21
                          $ 255 "AMR_PosTarget≔5"
                          global AMR_PosTarget=5
                        else:
                          $ 256 "ElseIf TASK.ID≟56"
                          if (TASK.ID == 56):
                            $ 257 "Task_info≔'Dose Powder'"
                            global Task_info="Dose Powder"
                            $ 258 "Parameters"
                            $ 259 "ITM_ID≔1"
                            global ITM_ID=1
                            $ 260 "target_weight≔(UGO.read_input('00','Target_weight'))/1000"
                            global target_weight=(UGO.read_input("00","Target_weight"))/1000
                            $ 261 "W_now≔(UGO.read_input('00','Container_weight'))/1000"
                            global W_now=(UGO.read_input("00","Container_weight"))/1000
                            $ 262 "Pow_name≔(UGO.read_input('00','Powder_name'))"
                            global Pow_name=(UGO.read_input("00","Powder_name"))
                            $ 263 "OBJ_Type≔6"
                            global OBJ_Type=6
                            $ 264 "JIG≔17"
                            global JIG=17
                            $ 265 "AMR_PosTarget≔5"
                            global AMR_PosTarget=5
                          else:
                            $ 266 "ElseIf TASK.ID≟57"
                            if (TASK.ID == 57):
                              $ 267 "Task_info≔'Recipe Powder dosing'"
                              global Task_info="Recipe Powder dosing"
                              $ 268 "Parameters"
                              $ 269 "ITM_ID≔1"
                              global ITM_ID=1
                              $ 270 "Pow_A≔(UGO.read_input('00','PowderA'))"
                              global Pow_A=(UGO.read_input("00","PowderA"))
                              $ 271 "Pow_B≔(UGO.read_input('00','PowderB'))"
                              global Pow_B=(UGO.read_input("00","PowderB"))
                              $ 272 "Pow_C≔(UGO.read_input('00','PowderC'))"
                              global Pow_C=(UGO.read_input("00","PowderC"))
                              $ 273 "Total_weight≔(UGO.read_input('00','Total_weight'))/1000"
                              global Total_weight=(UGO.read_input("00","Total_weight"))/1000
                              $ 274 "Pow_A_percent≔(UGO.read_input('00','PowderA_percentage'))/100"
                              global Pow_A_percent=(UGO.read_input("00","PowderA_percentage"))/100
                              $ 275 "Pow_B_percent≔(UGO.read_input('00','PowderB_percentage'))/100"
                              global Pow_B_percent=(UGO.read_input("00","PowderB_percentage"))/100
                              $ 276 "Pow_C_percent≔(UGO.read_input('00','PowderC_percentage'))/100"
                              global Pow_C_percent=(UGO.read_input("00","PowderC_percentage"))/100
                              $ 277 "OBJ_Type≔6"
                              global OBJ_Type=6
                              $ 278 "JIG≔17"
                              global JIG=17
                              $ 279 "AMR_PosTarget≔5"
                              global AMR_PosTarget=5
                            else:
                              $ 280 "ElseIf TASK.ID≟58"
                              if (TASK.ID == 58):
                                $ 281 "Task_info≔'Pick Powder containers'"
                                global Task_info="Pick Powder containers"
                                $ 282 "Parameters"
                                $ 283 "ITM_ID≔1"
                                global ITM_ID=1
                                $ 284 "OBJ_Type≔6"
                                global OBJ_Type=6
                                $ 285 "JIG≔15"
                                global JIG=15
                                $ 286 "AMR_PosTarget≔3"
                                global AMR_PosTarget=3
                              else:
                                $ 287 "ElseIf TASK.ID≟59"
                                if (TASK.ID == 59):
                                  $ 288 "Task_info≔'Empty Powder container'"
                                  global Task_info="Empty Powder container"
                                  $ 289 "Parameters"
                                  $ 290 "ITM_ID≔1"
                                  global ITM_ID=1
                                  $ 292 "Pow_name≔(UGO.read_input('00','Powder_name'))"
                                  global Pow_name=(UGO.read_input("00","Powder_name"))
                                  $ 294 "target_weight≔(aa_weight_cont-empty_weight_g)*1000"
                                  global target_weight=(aa_weight_cont-empty_weight_g)*1000
                                  $ 295 "W_now≔target_weight"
                                  global W_now=target_weight
                                  $ 296 "send_picking_info(Pow_name,target_weight)"
                                  send_picking_info(Pow_name,target_weight)
                                  $ 297 "w_dosed_total≔0"
                                  global w_dosed_total=0
                                  $ 298 "OBJ_Type≔6"
                                  global OBJ_Type=6
                                  $ 299 "JIG≔17"
                                  global JIG=17
                                  $ 300 "AMR_PosTarget≔5"
                                  global AMR_PosTarget=5
                                else:
                                  $ 301 "ElseIf TASK.ID≟61"
                                  if (TASK.ID == 61):
                                    $ 302 "Task_info≔'Weigh, Place & Decap'"
                                    global Task_info="Weigh, Place & Decap"
                                    $ 303 "Parameters"
                                    $ 304 "ITM_ID≔1"
                                    global ITM_ID=1
                                    $ 305 "OBJ_Type≔6"
                                    global OBJ_Type=6
                                    $ 306 "JIG≔21"
                                    global JIG=21
                                    $ 307 "AMR_PosTarget≔5"
                                    global AMR_PosTarget=5
                                  else:
                                    $ 308 "ElseIf TASK.ID≟62"
                                    if (TASK.ID == 62):
                                      $ 309 "Task_info≔'Dose Powder'"
                                      global Task_info="Dose Powder"
                                      $ 310 "Parameters"
                                      $ 311 "ITM_ID≔1"
                                      global ITM_ID=1
                                      $ 313 "W_now≔aa_weight_cont"
                                      global W_now=aa_weight_cont
                                      $ 314 "Pow_name≔(UGO.read_input('00','Powder_name'))"
                                      global Pow_name=(UGO.read_input("00","Powder_name"))
                                      $ 315 "target_weight≔(UGO.read_input('00','Target_weight'))/1000"
                                      global target_weight=(UGO.read_input("00","Target_weight"))/1000
                                      $ 317 "params_init()"
                                      params_init()
                                      $ 318 "send_picking_info(Pow_name,target_weight)"
                                      send_picking_info(Pow_name,target_weight)
                                      $ 319 "OBJ_Type≔6"
                                      global OBJ_Type=6
                                      $ 320 "JIG≔17"
                                      global JIG=17
                                      $ 321 "AMR_PosTarget≔5"
                                      global AMR_PosTarget=5
                                    else:
                                      $ 322 "Else" "noBreak"
                                      $ 323 "set_error(ERROR_WRONG_ORDER)"
                                      set_error(ERROR_WRONG_ORDER)
                                    end
                                  end
                                end
                              end
                            end
                          end
                        end
                      end
                    end
                  end
                end
              end
            end
          end
        end
      end
      $ 324 "test ugo"
      $ 325 "Wait: 0.2"
      sleep(0.2)
      $ 326 "ugo_update_outputs()"
      ugo_update_outputs()
      $ 327 "If starting() and AMR_Done"
      if (starting()  and  AMR_Done):
        $ 328 "log_message(Task_info, 'New Task: ')"
        log_message(Task_info, "New Task: ")
        $ 329 "log_message(to_str(TASK.ID), 'Task_ID: ')"
        log_message(to_str(TASK.ID), "Task_ID: ")
        $ 330 "do_transition(keep_rxry=OBJ_Picked)"
        do_transition(keep_rxry=OBJ_Picked)
        $ 331 "STATE≔6"
        global STATE=6
        $ 332 "ugo_update_outputs()"
        ugo_update_outputs()
      end
    elif (6 == switch_1):
      $ 333 "Case 6"
      $ 334 "Execute"
      $ 335 "STATE_Info≔'Execute'"
      global STATE_Info="Execute"
      $ 336 "If  not CMD_Hold and not CMD_Suspend"
      global thread_flag_336=0
      thread Thread_if_336():
        $ 337 "Switch PROCESS_Step"
        switch_2 = PROCESS_Step
        $ 338 "Case 0"
        if (0 == switch_2):
          $ 339 "PROCESS_Info≔'process control'"
          global PROCESS_Info="process control"
          $ 340 "log_process(PROCESS_Info)"
          log_process(PROCESS_Info)
          $ 341 "process control"
          $ 342 "If  not AMR_AtTarget"
          if (  not  AMR_AtTarget):
            $ 343 "PROCESS_Step≔1"
            global PROCESS_Step=1
          else:
            $ 344 "ElseIf (( not ITM_Prepared and  not WRK_Done) or (ITM_Prepared and WRK_Done))"
            if (((  not  ITM_Prepared  and    not  WRK_Done)  or  (ITM_Prepared  and  WRK_Done))):
              $ 345 "PROCESS_Step≔2"
              global PROCESS_Step=2
            else:
              $ 346 "ElseIf  not WRK_Done"
              if (  not  WRK_Done):
                $ 347 "PROCESS_Step≔3"
                global PROCESS_Step=3
              else:
                $ 348 "Else" "noBreak"
                $ 349 "task finished"
                $ 350 "PROCESS_Info≔''"
                global PROCESS_Info=""
                $ 351 "STATE≔7"
                global STATE=7
                $ 352 "ugo_update_outputs()"
                ugo_update_outputs()
              end
            end
          end
        elif (1 == switch_2):
          $ 353 "Case 1"
          $ 354 "navigate"
          $ 355 "'MOVING THE uML'"
          # 'MOVING THE uML'
          $ 356 "PROCESS_Info≔'move to target'"
          global PROCESS_Info="move to target"
          $ 357 "log_process(PROCESS_Info)"
          log_process(PROCESS_Info)
          $ 358 "If TASK.ID≟1"
          if (TASK.ID == 1):
            $ 359 "Action≔51"
            global Action=51
          else:
            $ 360 "Else" "noBreak"
            $ 361 "Action≔52"
            global Action=52
          end
          $ 362 "Call Sub_AMR_MiR_V3"
          Sub_AMR_MiR_V3()
          $ 363 "If AMR_Done"
          if (AMR_Done):
            $ 364 "PROCESS_Step≔0"
            global PROCESS_Step=0
          end
        elif (2 == switch_2):
          $ 365 "Case 2"
          $ 366 "prepare"
          $ 367 "'THINGS THAT HAVE TO BE DONE ONCE IN A SEQUENCE,WORKFLOW'"
          # 'THINGS THAT HAVE TO BE DONE ONCE IN A SEQUENCE,WORKFLOW'
          $ 368 "PROCESS_Info≔'prepare for work'"
          global PROCESS_Info="prepare for work"
          $ 369 "log_process(PROCESS_Info)"
          log_process(PROCESS_Info)
          $ 370 "If TASK.WORK.ITM_ID_Src>1"
          if (TASK.WORK.ITM_ID_Src>1):
            $ 371 "ITM_ID≔TASK.WORK.ITM_ID_Src"
            global ITM_ID=TASK.WORK.ITM_ID_Src
          else:
            $ 372 "ElseIf TASK.WORK.ITM_ID_Tgt>1"
            if (TASK.WORK.ITM_ID_Tgt>1):
              $ 373 "ITM_ID≔TASK.WORK.ITM_ID_Tgt"
              global ITM_ID=TASK.WORK.ITM_ID_Tgt
            end
          end
          $ 374 "If  not ARM_Referenced and (ITM_ID≠0)"
          if (  not  ARM_Referenced  and  (ITM_ID != 0)):
            $ 375 "STP≔1"
            global STP=1
          else:
            $ 376 "ElseIf ARM_Referenced or (ITM_ID≟0)"
            if (ARM_Referenced  or  (ITM_ID == 0)):
              $ 377 "STP≔2"
              global STP=2
            end
          end
          $ 378 "Switch STP"
          switch_3 = STP
          $ 379 "Case 1"
          if (1 == switch_3):
            $ 380 "reference"
            $ 381 "STP_Info≔'reference at target position'"
            global STP_Info="reference at target position"
            $ 382 "log_step(STP_Info)"
            log_step(STP_Info)
            $ 383 "If ITM_ID≟1"
            if (ITM_ID == 1):
              $ 384 "CAM_Done≔ True "
              global CAM_Done=  True
            else:
              $ 385 "Else" "noBreak"
              $ 386 "Action≔131"
              global Action=131
              $ 387 "Call Sub_Vision_V18"
              Sub_Vision_V18()
            end
            $ 389 "If CAM_Done and  not ERROR.FLAG"
            if (CAM_Done  and    not  ERROR.FLAG):
              $ 390 "log_step('ARM referenced')"
              log_step("ARM referenced")
              $ 391 "ARM_Referenced≔ True "
              global ARM_Referenced=  True
            end
          elif (2 == switch_3):
            $ 392 "Case 2"
            $ 393 "manipulate"
            $ 394 "STP_Info≔'manipulate item'"
            global STP_Info="manipulate item"
            $ 395 "log_step(STP_Info)"
            log_step(STP_Info)
            $ 396 "'In case pressing button is needed'"
            # 'In case pressing button is needed'
            $ 397 "If found_in_list(ITM_ID, ITM_ID_List)"
            if (found_in_list(ITM_ID, ITM_ID_List)):
              $ 398 "Switch ITM_ID"
              switch_4 = ITM_ID
              $ 399 "Case 0"
              if (0 == switch_4):
                $ 400 "ITM_Manipulated≔ not ITM_Manipulated"
                global ITM_Manipulated=  not  ITM_Manipulated
              elif (1 == switch_4):
                $ 401 "Case 1"
                $ 402 "ITM_Manipulated≔ not ITM_Manipulated"
                global ITM_Manipulated=  not  ITM_Manipulated
              elif (2 == switch_4):
                $ 403 "Case 2"
              else:
                $ 413 "Default Case"
                $ 414 "ITM_Manipulated≔ not ITM_Manipulated"
                global ITM_Manipulated=  not  ITM_Manipulated
              end
            end
          end
          $ 415 "ITM_Prepared≔(ITM_Manipulated or  not found_in_list(ITM_ID, ITM_ID_List)) and (ARM_Referenced or ITM_ID≟0) and  not WRK_Done"
          global ITM_Prepared=(ITM_Manipulated  or    not  found_in_list(ITM_ID, ITM_ID_List))  and  (ARM_Referenced  or  ITM_ID == 0)  and    not  WRK_Done
          $ 416 "STP≔0"
          global STP=0
          $ 417 "STP_Info≔''"
          global STP_Info=""
          $ 418 "PROCESS_Step≔0"
          global PROCESS_Step=0
        elif (3 == switch_2):
          $ 419 "Case 3"
          $ 420 "work"
          $ 421 "'ADD EVERY MACHINE, OBJECT, STATION TO WORK ON'"
          # 'ADD EVERY MACHINE, OBJECT, STATION TO WORK ON'
          $ 422 "Switch ITM_ID"
          switch_3 = ITM_ID
          $ 423 "Case 1"
          if (1 == switch_3):
            $ 424 "uLM"
            $ 425 "If TASK.ID≟12"
            if (TASK.ID == 12):
              $ 426 "fill racks"
              $ 427 "Action≔151"
              global Action=151
              $ 428 "Call Sub_Vision_V18"
              Sub_Vision_V18()
              $ 429 "If  not ERROR.FLAG"
              if (  not  ERROR.FLAG):
                $ 430 "Actions for the task"
                $ 431 "Action≔1"
                global Action=1
                $ 432 "JIG≔2"
                global JIG=2
                $ 433 "JIG_Slot≔CAM_Result[0]"
                global JIG_Slot=CAM_Result[0]
                $ 434 "OBJ_Nbr≔CAM_Result[0]"
                global OBJ_Nbr=CAM_Result[0]
                $ 435 "OBJ_Type≔2"
                global OBJ_Type=2
                $ 436 "Call Sub_Action_V4"
                Sub_Action_V4()
                $ 437 "If OBJ_Picked"
                if (OBJ_Picked):
                  $ 438 "CAM_Result.remove(0)"
                  CAM_Result.remove(0)
                  $ 439 "PRC_TubCounter≔PRC_TubCounter+1"
                  global PRC_TubCounter=PRC_TubCounter+1
                  $ 440 "If PRC_TubCounter%4≟0"
                  if (PRC_TubCounter%4 == 0):
                    $ 441 "JIG_Slot≔4"
                    global JIG_Slot=4
                  else:
                    $ 442 "Else" "noBreak"
                    $ 443 "JIG_Slot≔PRC_TubCounter%4"
                    global JIG_Slot=PRC_TubCounter%4
                  end
                  $ 444 "OBJ_Nbr≔ceil(PRC_TubCounter/4)"
                  global OBJ_Nbr=ceil(PRC_TubCounter/4)
                  $ 445 "Action≔2"
                  global Action=2
                  $ 446 "JIG≔4"
                  global JIG=4
                  $ 447 "Call Sub_Action_V4"
                  Sub_Action_V4()
                  $ 448 "Action≔151"
                  global Action=151
                  $ 449 "Call Sub_Vision_V18"
                  Sub_Vision_V18()
                end
              end
              $ 450 "If (CAM_Captures≥CAM_PRM_Retries) or (PRC_TubCounter≥32)"
              if ((CAM_Captures >= CAM_PRM_Retries)  or  (PRC_TubCounter >= 32)):
                $ 451 "PROCESS_Step≔0"
                global PROCESS_Step=0
                $ 452 "WRK_Done≔ True "
                global WRK_Done=  True
              end
            else:
              $ 453 "ElseIf TASK.ID≟13"
              if (TASK.ID == 13):
                $ 454 "Dose Powder"
                $ 455 "Action≔131"
                global Action=131
                $ 456 "Call Sub_Vision_V18"
                Sub_Vision_V18()
                $ 457 "Action≔34"
                global Action=34
                $ 458 "Call Sub_Action_V4"
                Sub_Action_V4()
                $ 459 "PROCESS_Step≔0"
                global PROCESS_Step=0
                $ 460 "WRK_Done≔ True "
                global WRK_Done=  True
              else:
                $ 461 "ElseIf TASK.ID≟49"
                if (TASK.ID == 49):
                  $ 462 "Pick Powder container"
                  $ 463 "Action≔131"
                  global Action=131
                  $ 464 "Call Sub_Vision_V18"
                  Sub_Vision_V18()
                  $ 465 "Action≔35"
                  global Action=35
                  $ 466 "Call Sub_Action_V4"
                  Sub_Action_V4()
                  $ 467 "PROCESS_Step≔0"
                  global PROCESS_Step=0
                  $ 468 "WRK_Done≔ True "
                  global WRK_Done=  True
                else:
                  $ 469 "ElseIf TASK.ID≟50"
                  if (TASK.ID == 50):
                    $ 470 "Decap containers"
                    $ 471 "Action≔36"
                    global Action=36
                    $ 472 "Call Sub_Action_V4"
                    Sub_Action_V4()
                    $ 473 "PROCESS_Step≔0"
                    global PROCESS_Step=0
                    $ 474 "WRK_Done≔ True "
                    global WRK_Done=  True
                  else:
                    $ 475 "ElseIf TASK.ID≟51"
                    if (TASK.ID == 51):
                      $ 476 "Detect Spatula and transfer powder"
                      $ 477 "Action≔131"
                      global Action=131
                      $ 478 "Call Sub_Vision_V18"
                      Sub_Vision_V18()
                      $ 479 "Action≔37"
                      global Action=37
                      $ 480 "Call Sub_Action_V4"
                      Sub_Action_V4()
                      $ 481 "PROCESS_Step≔0"
                      global PROCESS_Step=0
                      $ 482 "WRK_Done≔ True "
                      global WRK_Done=  True
                    else:
                      $ 483 "ElseIf TASK.ID≟52"
                      if (TASK.ID == 52):
                        $ 484 "Pick Powder container"
                        $ 485 "Action≔131"
                        global Action=131
                        $ 486 "Call Sub_Vision_V18"
                        Sub_Vision_V18()
                        $ 487 "Action≔39"
                        global Action=39
                        $ 488 "Call Sub_Action_V4"
                        Sub_Action_V4()
                        $ 489 "PROCESS_Step≔0"
                        global PROCESS_Step=0
                        $ 490 "WRK_Done≔ True "
                        global WRK_Done=  True
                      else:
                        $ 491 "ElseIf TASK.ID≟53"
                        if (TASK.ID == 53):
                          $ 492 "Decap containerA"
                          $ 493 "Action≔40"
                          global Action=40
                          $ 494 "Call Sub_Action_V4"
                          Sub_Action_V4()
                          $ 495 "PROCESS_Step≔0"
                          global PROCESS_Step=0
                          $ 496 "WRK_Done≔ True "
                          global WRK_Done=  True
                        else:
                          $ 497 "ElseIf TASK.ID≟55"
                          if (TASK.ID == 55):
                            $ 498 "Place Powder"
                            $ 499 "Action≔131"
                            global Action=131
                            $ 500 "Call Sub_Vision_V18"
                            Sub_Vision_V18()
                            $ 501 "Action≔41"
                            global Action=41
                            $ 502 "Call Sub_Action_V4"
                            Sub_Action_V4()
                            $ 503 "PROCESS_Step≔0"
                            global PROCESS_Step=0
                            $ 504 "WRK_Done≔ True "
                            global WRK_Done=  True
                          else:
                            $ 505 "ElseIf TASK.ID≟54"
                            if (TASK.ID == 54):
                              $ 506 "Empty and swap container"
                              $ 507 "Action≔131"
                              global Action=131
                              $ 508 "Call Sub_Vision_V18"
                              Sub_Vision_V18()
                              $ 509 "Action≔42"
                              global Action=42
                              $ 510 "Call Sub_Action_V4"
                              Sub_Action_V4()
                              $ 511 "PROCESS_Step≔0"
                              global PROCESS_Step=0
                              $ 512 "WRK_Done≔ True "
                              global WRK_Done=  True
                            else:
                              $ 513 "ElseIf TASK.ID≟56"
                              if (TASK.ID == 56):
                                $ 514 "Dispense Powder"
                                $ 515 "Action≔131"
                                global Action=131
                                $ 516 "Call Sub_Vision_V18"
                                Sub_Vision_V18()
                                $ 517 "Action≔43"
                                global Action=43
                                $ 518 "Call Sub_Action_V4"
                                Sub_Action_V4()
                                $ 519 "PROCESS_Step≔0"
                                global PROCESS_Step=0
                                $ 520 "WRK_Done≔ True "
                                global WRK_Done=  True
                              else:
                                $ 521 "ElseIf TASK.ID≟57"
                                if (TASK.ID == 57):
                                  $ 522 "Recipe Dosing"
                                  $ 523 "Action≔48"
                                  global Action=48
                                  $ 524 "Call Sub_Action_V4"
                                  Sub_Action_V4()
                                  $ 541 "PROCESS_Step≔0"
                                  global PROCESS_Step=0
                                  $ 542 "WRK_Done≔ True "
                                  global WRK_Done=  True
                                else:
                                  $ 543 "ElseIf TASK.ID≟58"
                                  if (TASK.ID == 58):
                                    $ 544 "Pick Powder containers"
                                    $ 545 "Num_cont_picked≔0"
                                    global Num_cont_picked=0
                                    $ 546 "powder_position≔'Position1'"
                                    global powder_position="Position1"
                                    $ 547 "Loop Num_cont_picked<3"
                                    while (Num_cont_picked<3):
                                      $ 548 "Action≔131"
                                      global Action=131
                                      $ 549 "Call Sub_Vision_V18"
                                      Sub_Vision_V18()
                                      $ 550 "Action≔47"
                                      global Action=47
                                      $ 551 "Call Sub_Action_V4"
                                      Sub_Action_V4()
                                    end
                                    $ 552 "PROCESS_Step≔0"
                                    global PROCESS_Step=0
                                    $ 553 "WRK_Done≔ True "
                                    global WRK_Done=  True
                                  else:
                                    $ 554 "ElseIf TASK.ID≟59"
                                    if (TASK.ID == 59):
                                      $ 555 "Empty powder container"
                                      $ 556 "Action≔131"
                                      global Action=131
                                      $ 557 "Call Sub_Vision_V18"
                                      Sub_Vision_V18()
                                      $ 558 "Action≔50"
                                      global Action=50
                                      $ 559 "Call Sub_Action_V4"
                                      Sub_Action_V4()
                                      $ 560 "PROCESS_Step≔0"
                                      global PROCESS_Step=0
                                      $ 561 "WRK_Done≔ True "
                                      global WRK_Done=  True
                                    else:
                                      $ 562 "ElseIf TASK.ID≟61"
                                      if (TASK.ID == 61):
                                        $ 563 "Place Powder"
                                        $ 564 "Action≔131"
                                        global Action=131
                                        $ 565 "Call Sub_Vision_V18"
                                        Sub_Vision_V18()
                                        $ 566 "Action≔51"
                                        global Action=51
                                        $ 567 "Call Sub_Action_V4"
                                        Sub_Action_V4()
                                        $ 568 "PROCESS_Step≔0"
                                        global PROCESS_Step=0
                                        $ 569 "WRK_Done≔ True "
                                        global WRK_Done=  True
                                      else:
                                        $ 570 "ElseIf TASK.ID≟62"
                                        if (TASK.ID == 62):
                                          $ 571 "Dose Powder"
                                          $ 572 "Action≔131"
                                          global Action=131
                                          $ 573 "Call Sub_Vision_V18"
                                          Sub_Vision_V18()
                                          $ 574 "Action≔52"
                                          global Action=52
                                          $ 575 "Call Sub_Action_V4"
                                          Sub_Action_V4()
                                          $ 576 "PROCESS_Step≔0"
                                          global PROCESS_Step=0
                                          $ 577 "WRK_Done≔ True "
                                          global WRK_Done=  True
                                        end
                                      end
                                    end
                                  end
                                end
                              end
                            end
                          end
                        end
                      end
                    end
                  end
                end
              end
            end
          elif (2 == switch_3):
            $ 578 "Case 2"
          elif (5 == switch_3):
            $ 620 "Case 5"
          elif (20 == switch_3):
            $ 628 "Case 20"
          elif (43 == switch_3):
            $ 690 "Case 43"
          else:
            $ 698 "Default Case"
            $ 699 "WRK_Done≔ True "
            global WRK_Done=  True
            $ 700 "PROCESS_Step≔0"
            global PROCESS_Step=0
          end
        end
        thread_flag_336 = 1
      end
      if (  not  CMD_Hold and not CMD_Suspend):
        global thread_handler_336=run Thread_if_336()
        while (thread_flag_336 == 0):
          if not(  not  CMD_Hold and not CMD_Suspend):
            kill thread_handler_336
            thread_flag_336 = 2
          else:
            sync()
          end
        end
      else:
        thread_flag_336 = 2
      end
      $ 701 "If CMD_Hold"
      if (CMD_Hold):
        $ 702 "STATE≔9"
        global STATE=9
        $ 703 "ugo_update_outputs()"
        ugo_update_outputs()
      else:
        $ 704 "ElseIf CMD_Suspend"
        if (CMD_Suspend):
          $ 705 "STATE≔12"
          global STATE=12
          $ 706 "ugo_update_outputs()"
          ugo_update_outputs()
        end
      end
    elif (7 == switch_1):
      $ 707 "Case 7"
      $ 708 "Completing"
      $ 709 "STATE_Info≔'Completing'"
      global STATE_Info="Completing"
      $ 710 "'ADD COMMANDS FOR COMPLETING THE PROCESS'"
      # 'ADD COMMANDS FOR COMPLETING THE PROCESS'
      $ 711 "do_transition(keep_rxry=OBJ_Picked)"
      do_transition(keep_rxry=OBJ_Picked)
      $ 712 "Call Sub_AMR_MiR_V3"
      Sub_AMR_MiR_V3()
      $ 713 "If completing() and AMR_Done"
      if (completing()  and  AMR_Done):
        $ 714 "STATE≔8"
        global STATE=8
        $ 715 "ugo_update_outputs()"
        ugo_update_outputs()
      end
    elif (8 == switch_1):
      $ 716 "Case 8"
      $ 717 "Complete"
      $ 718 "STATE_Info≔'Complete'"
      global STATE_Info="Complete"
      $ 719 "If CMD_Reset"
      if (CMD_Reset):
        $ 720 "STATE≔3"
        global STATE=3
        $ 721 "ugo_update_outputs()"
        ugo_update_outputs()
      end
    elif (9 == switch_1):
      $ 722 "Case 9"
      $ 723 "Holding"
      $ 724 "STATE_Info≔'Holding'"
      global STATE_Info="Holding"
      $ 725 "stopl(0.5)"
      stopl(0.5)
      $ 726 "Call Sub_AMR_MiR_V3"
      Sub_AMR_MiR_V3()
      $ 727 "If holding() and AMR_Done"
      if (holding()  and  AMR_Done):
        $ 728 "STATE≔10"
        global STATE=10
        $ 729 "ugo_update_outputs()"
        ugo_update_outputs()
      end
    elif (10 == switch_1):
      $ 730 "Case 10"
      $ 731 "Held"
      $ 732 "STATE_Info≔'Held'"
      global STATE_Info="Held"
      $ 733 "If CMD_Unhold"
      if (CMD_Unhold):
        $ 734 "end_freedrive_mode()"
        end_freedrive_mode()
        $ 735 "STATE≔11"
        global STATE=11
        $ 736 "ugo_update_outputs()"
        ugo_update_outputs()
      else:
        $ 737 "ElseIf FNC_Freedrive"
        if (FNC_Freedrive):
          $ 738 "freedrive_mode()"
          freedrive_mode()
        else:
          $ 739 "Else" "noBreak"
          $ 740 "end_freedrive_mode()"
          end_freedrive_mode()
        end
      end
    elif (11 == switch_1):
      $ 741 "Case 11"
      $ 742 "Unholding"
      $ 743 "STATE_Info≔'Unholding'"
      global STATE_Info="Unholding"
      $ 744 "Clearing"
      $ 745 "Switch ERROR.ID"
      switch_2 = ERROR.ID
      $ 746 "Case 1002"
      if (1002 == switch_2):
        $ 747 "AMR_AtTarget≔ False "
        global AMR_AtTarget=  False
        $ 748 "ARM_Referenced≔ False "
        global ARM_Referenced=  False
        $ 749 "ITM_Prepared≔ False "
        global ITM_Prepared=  False
        $ 750 "PROCESS_Step≔1"
        global PROCESS_Step=1
      elif (2007 == switch_2):
        $ 751 "Case 2007"
        $ 752 "PROCESS_Step≔1"
        global PROCESS_Step=1
      end
      $ 753 "reset_error()"
      reset_error()
      $ 754 "reset_warning()"
      reset_warning()
      $ 755 "OBJ_Picked≔gripper_has_object()"
      global OBJ_Picked=gripper_has_object()
      $ 756 "Call Sub_AMR_MiR_V3"
      Sub_AMR_MiR_V3()
      $ 757 "If unholding() and AMR_Done"
      if (unholding()  and  AMR_Done):
        $ 758 "STATE≔6"
        global STATE=6
        $ 759 "ugo_update_outputs()"
        ugo_update_outputs()
      end
    elif (12 == switch_1):
      $ 760 "Case 12"
      $ 761 "Suspending"
      $ 762 "STATE_Info≔'Suspending'"
      global STATE_Info="Suspending"
      $ 763 "PROCESS_Info≔str_cat(PROCESS_Info, ' suspended')"
      global PROCESS_Info=str_cat(PROCESS_Info, " suspended")
      $ 764 "If suspending()"
      if (suspending()):
        $ 765 "STATE≔13"
        global STATE=13
        $ 766 "ugo_update_outputs()"
        ugo_update_outputs()
      end
    elif (13 == switch_1):
      $ 767 "Case 13"
      $ 768 "Suspended"
      $ 769 "STATE_Info≔'Suspended'"
      global STATE_Info="Suspended"
      $ 770 "Call Sub_AMR_MiR_V3"
      Sub_AMR_MiR_V3()
      $ 771 "If CMD_Unsuspend"
      if (CMD_Unsuspend):
        $ 772 "STATE≔14"
        global STATE=14
        $ 773 "ugo_update_outputs()"
        ugo_update_outputs()
      end
    elif (14 == switch_1):
      $ 774 "Case 14"
      $ 775 "Unsuspending"
      $ 776 "STATE_Info≔'Unsuspending'"
      global STATE_Info="Unsuspending"
      $ 777 "PROCESS_Step≔0"
      global PROCESS_Step=0
      $ 778 "If unsuspending()"
      if (unsuspending()):
        $ 779 "STATE≔6"
        global STATE=6
        $ 780 "ugo_update_outputs()"
        ugo_update_outputs()
      end
    elif (15 == switch_1):
      $ 781 "Case 15"
      $ 782 "Aborting"
      $ 783 "STATE_Info≔'Aborting'"
      global STATE_Info="Aborting"
      $ 784 "If aborting()"
      if (aborting()):
        $ 785 "STATE≔16"
        global STATE=16
        $ 786 "ugo_update_outputs()"
        ugo_update_outputs()
      end
    elif (16 == switch_1):
      $ 787 "Case 16"
      $ 788 "Aborted"
      $ 789 "STATE_Info≔'Aborted'"
      global STATE_Info="Aborted"
      $ 790 "If CMD_Clear"
      if (CMD_Clear):
        $ 791 "STATE≔17"
        global STATE=17
        $ 792 "ugo_update_outputs()"
        ugo_update_outputs()
      end
    elif (17 == switch_1):
      $ 793 "Case 17"
      $ 794 "Clearing"
      $ 795 "STATE_Info≔'Clearing'"
      global STATE_Info="Clearing"
      $ 796 "Clearing"
      $ 797 "reset_warning()"
      reset_warning()
      $ 798 "reset_error()"
      reset_error()
      $ 799 "If clearing()"
      if (clearing()):
        $ 800 "STATE≔2"
        global STATE=2
        $ 801 "ugo_update_outputs()"
        ugo_update_outputs()
      end
    end
    $ 802 "log_state(STATE_Info)"
    log_state(STATE_Info)
    $ 803 "log_warning(WARNING.MSG)"
    log_warning(WARNING.MSG)
    $ 804 "log_error(ERROR.MSG)"
    log_error(ERROR.MSG)
    $ 805 "Times"
    $ 806 "Switch STATE"
    switch_1 = STATE
    $ 807 "Case 1"
    if (1 == switch_1):
      $ 808 "TM_St_Stopping≔get_time(STATE_Times[STATE-1])"
      global TM_St_Stopping=get_time(STATE_Times[STATE-1])
    elif (2 == switch_1):
      $ 809 "Case 2"
      $ 810 "TM_St_Stopped≔get_time(STATE_Times[STATE-1])"
      global TM_St_Stopped=get_time(STATE_Times[STATE-1])
    elif (3 == switch_1):
      $ 811 "Case 3"
      $ 812 "TM_St_Resetting≔get_time(STATE_Times[STATE-1])"
      global TM_St_Resetting=get_time(STATE_Times[STATE-1])
    elif (4 == switch_1):
      $ 813 "Case 4"
      $ 814 "TM_St_Idle≔get_time(STATE_Times[STATE-1])"
      global TM_St_Idle=get_time(STATE_Times[STATE-1])
    elif (5 == switch_1):
      $ 815 "Case 5"
      $ 816 "TM_St_Starting≔get_time(STATE_Times[STATE-1])"
      global TM_St_Starting=get_time(STATE_Times[STATE-1])
    elif (6 == switch_1):
      $ 817 "Case 6"
      $ 818 "TM_St_Execute≔get_time(STATE_Times[STATE-1])"
      global TM_St_Execute=get_time(STATE_Times[STATE-1])
    elif (7 == switch_1):
      $ 819 "Case 7"
      $ 820 "TM_St_Completin≔get_time(STATE_Times[STATE-1])"
      global TM_St_Completin=get_time(STATE_Times[STATE-1])
    elif (8 == switch_1):
      $ 821 "Case 8"
      $ 822 "TM_St_Complete≔get_time(STATE_Times[STATE-1])"
      global TM_St_Complete=get_time(STATE_Times[STATE-1])
    elif (9 == switch_1):
      $ 823 "Case 9"
      $ 824 "TM_St_Holding≔get_time(STATE_Times[STATE-1])"
      global TM_St_Holding=get_time(STATE_Times[STATE-1])
    elif (10 == switch_1):
      $ 825 "Case 10"
      $ 826 "TM_St_Held≔get_time(STATE_Times[STATE-1])"
      global TM_St_Held=get_time(STATE_Times[STATE-1])
    elif (11 == switch_1):
      $ 827 "Case 11"
      $ 828 "TM_St_Unholding≔get_time(STATE_Times[STATE-1])"
      global TM_St_Unholding=get_time(STATE_Times[STATE-1])
    elif (12 == switch_1):
      $ 829 "Case 12"
      $ 830 "TM_St_Suspendin≔get_time(STATE_Times[STATE-1])"
      global TM_St_Suspendin=get_time(STATE_Times[STATE-1])
    elif (13 == switch_1):
      $ 831 "Case 13"
      $ 832 "TM_St_Suspended≔get_time(STATE_Times[STATE-1])"
      global TM_St_Suspended=get_time(STATE_Times[STATE-1])
    elif (14 == switch_1):
      $ 833 "Case 14"
      $ 834 "TM_St_Unsuspend≔get_time(STATE_Times[STATE-1])"
      global TM_St_Unsuspend=get_time(STATE_Times[STATE-1])
    elif (15 == switch_1):
      $ 835 "Case 15"
      $ 836 "TM_St_Aborting≔get_time(STATE_Times[STATE-1])"
      global TM_St_Aborting=get_time(STATE_Times[STATE-1])
    elif (16 == switch_1):
      $ 837 "Case 16"
      $ 838 "TM_St_Aborted≔get_time(STATE_Times[STATE-1])"
      global TM_St_Aborted=get_time(STATE_Times[STATE-1])
    elif (17 == switch_1):
      $ 839 "Case 17"
      $ 840 "TM_St_Clearing≔get_time(STATE_Times[STATE-1])"
      global TM_St_Clearing=get_time(STATE_Times[STATE-1])
    end
    $ 842 "Wait: 0.1"
    sleep(0.1)
  end
end
